Fanuc KAREL source: KT00589.KL

PROGRAM KT00589
%NOLOCKGROUP
VAR
  S1: STRING[80]
  S2: STRING[80]
  OUT: STRING[80]
BEGIN
  S1 = 'A'
  S2 = 'B'
  S1 = 'A'
  S2 = 'B'
  OUT = S1 + S2
END KT00589
